DATA_BLOCK "Current_state_of_Bay0"
{ S7_Optimized_Access := 'TRUE' }
VERSION : 0.1
NON_RETAIN
   VAR
      Bay0 : Array[0..3, 0..11] of UInt;
   END_VAR


BEGIN
   Bay0[0,0] := 101;
   Bay0[0,1] := 0;
   Bay0[0,2] := 0;
   Bay0[0,3] := 0;
   Bay0[0,4] := 0;
   Bay0[0,5] := 0;
   Bay0[0,6] := 0;
   Bay0[0,7] := 0;
   Bay0[0,8] := 0;
   Bay0[0,9] := 0;
   Bay0[0,10] := 0;
   Bay0[0,11] := 0;
   Bay0[1,0] := 102;
   Bay0[1,1] := 0;
   Bay0[1,2] := 0;
   Bay0[1,3] := 0;
   Bay0[1,4] := 0;
   Bay0[1,5] := 0;
   Bay0[1,6] := 0;
   Bay0[1,7] := 0;
   Bay0[1,8] := 0;
   Bay0[1,9] := 0;
   Bay0[1,10] := 0;
   Bay0[1,11] := 0;
   Bay0[2,0] := 103;
   Bay0[2,1] := 0;
   Bay0[2,2] := 0;
   Bay0[2,3] := 0;
   Bay0[2,4] := 0;
   Bay0[2,5] := 0;
   Bay0[2,6] := 0;
   Bay0[2,7] := 0;
   Bay0[2,8] := 0;
   Bay0[2,9] := 0;
   Bay0[2,10] := 0;
   Bay0[2,11] := 0;
   Bay0[3,0] := 104;
   Bay0[3,1] := 0;
   Bay0[3,2] := 0;
   Bay0[3,3] := 0;
   Bay0[3,4] := 0;
   Bay0[3,5] := 0;
   Bay0[3,6] := 0;
   Bay0[3,7] := 0;
   Bay0[3,8] := 0;
   Bay0[3,9] := 0;
   Bay0[3,10] := 0;
   Bay0[3,11] := 0;

END_DATA_BLOCK

